// TIA Portal V21 export
// export: Created 2026-11-10T07:02:24.4553878Z, ExportSetting WithDefaults, DisplayName Totally Integrated Automation Portal, DisplayVersion V21 Update 3, DisplayName STEP 7 Professional, DisplayVersion V21 Update 3, DisplayName STEP 7 Safety, DisplayVersion V21, DisplayName Tech WebApplication, DisplayVersion V21, DisplayName WinCC Basic/Comfort/Advanced, DisplayVersion V21 Update 3, DisplayName WinCC Unified, DisplayVersion V21 Update 3
FUNCTION "FC_SclMath" : Void   // FC7, SCL
{ S7_Optimized_Access := 'TRUE' }
VERSION : 0.1
// stored: AutoNumber true, IsIECCheckEnabled false, SetENOAutomatically false, UDAEnableTagReadback false
   VAR_TEMP
      i : Int;
      j : Int;
      d : DInt;
      r : Real;
      r2 : Real;
      lr : LReal;
      "b" : Bool;
      w : Word;
      dw : DWord;
      "by" : Byte;
      t : Time;
   END_VAR
BEGIN
   #r := ABS(#r2);
   #r := SQRT(#r2);
   #r := SQR(#r2);
   #r := LN(#r2);
   #r := EXP(#r2);
   #r := SIN(#r2);
   #r := COS(#r2);
   #r := TAN(#r2);
   #r := ASIN(#r2);
   #r := ACOS(#r2);
   #r := ATAN(#r2);
   #i := ABS(#j);
   #i := MIN(IN1 := #i, IN2 := #j);
   #i := MAX(IN1 := #i, IN2 := #j);
   #i := LIMIT(MN := 0, IN := #i, MX := 100);
   #i := MIN(IN1 := #i, IN2 := #j, IN3 := 5);
   #i := MAX(IN1 := #i, IN2 := #j, IN3 := 5);
   #i := SEL(G := #b, IN0 := #i, IN1 := #j);
   #i := MUX(K := #j, IN0 := 1, IN1 := 2, IN2 := 3);
   #r := INT_TO_REAL(#i);
   #i := REAL_TO_INT(#r);
   #d := REAL_TO_DINT(#r);
   #i := DINT_TO_INT(#d);
   #d := INT_TO_DINT(#i);
   #d := TRUNC(#r);
   #d := ROUND(#r);
   #d := CEIL(#r);
   #d := FLOOR(#r);
   #r := DINT_TO_REAL(#d);
   #w := INT_TO_WORD(#i);
   #i := WORD_TO_INT(#w);
   #dw := SHL(IN := #dw, N := 2);
   #dw := SHR(IN := #dw, N := 2);
   #dw := ROL(IN := #dw, N := 1);
   #dw := ROR(IN := #dw, N := 1);
   #w := SHL(IN := #w, N := 1);
   #by := BYTE#16#01;
   #t := INT_TO_TIME(#i);
   #r := NORM_X(MIN := 0, VALUE := #i, MAX := 27648);
   #i := SCALE_X(MIN := 0, VALUE := #r, MAX := 27648);
   #d := DWORD_TO_DINT(#dw);
   #dw := DINT_TO_DWORD(#d);
   #r := FRAC(#r2);
END_FUNCTION
